(* IEC 61131-3 sources: plc-vscode/tests/st/test-ready/rusty/tests/lit/single/builtin, 5 files *)

(* ---- adr_ptr_arith_runtime.st ---- *)
// RUN: (%COMPILE %s && %RUN) | %CHECK %s
//
// `ADR(x) + N` is byte-stride pointer arithmetic — `ADR` is declared to
// return LWORD, so the `+` flows through the integer-arithmetic path; the
// receiver pointer ends up `N` bytes past the operand. Regression for #1749
// (previously panicked in `create_llvm_int_binary_expression`).

FUNCTION main
VAR
    arr : ARRAY[0..7] OF BYTE := [0, 0, 0, 0, 0, 0, 0, 0];
    pt  : REF_TO BYTE;
END_VAR

pt := ADR(arr) + 4;
pt^ := BYTE#16#AB;

// CHECK: arr[4]=171
printf('arr[4]=%d$N', arr[4]);

pt := ADR(arr) + 7;
pt^ := BYTE#16#5C;

// CHECK: arr[7]=92
printf('arr[7]=%d$N', arr[7]);

// Subtraction flows through the same path: take a pointer past the end
// and walk back. Writing to arr[2] via `ADR(arr[6]) - 4`.
pt := ADR(arr[6]) - 4;
pt^ := BYTE#16#11;

// CHECK: arr[2]=17
printf('arr[2]=%d$N', arr[2]);
END_FUNCTION

(* ---- shl_and_shr_must_cast_left_and_right_correctly.st ---- *)
// RUN: (%COMPILE %s && %RUN) | %CHECK %s

// SHL and SHR must cast left and right correctly
FUNCTION main
VAR
    value : BYTE;
END_VAR

value := BIT_LOAD_B2(BYTE#255, TRUE, 2, 2);

// CHECK: 255
printf('%d$N', value);

value := BIT_LOAD_B2(BYTE#255, FALSE, 2, 2);

// CHECK: 243
printf('%d$N', value);

END_FUNCTION

FUNCTION BIT_LOAD_B2 : BYTE
VAR_INPUT
	I : BYTE;
	D : BOOL;
	P : INT;
	N : INT;
END_VAR
VAR
    result : BYTE;
END_VAR

IF D THEN
	BIT_LOAD_B2 := ROL(SHR(BYTE#255, 8 - N) OR ROR(I, P), P);
ELSE
	BIT_LOAD_B2 := ROL(SHL(BYTE#255, N) AND ROR(I, P), P);
END_IF;

END_FUNCTION

(* ---- shl_must_be_usable_with_integers.st ---- *)
// RUN: (%COMPILE %s && %RUN) | %CHECK %s

// SHL must be usable with integers
FUNCTION main
VAR
    a : INT;
END_VAR
a := SHL(21,2);

// CHECK: 84
printf('%d$N', a);
END_FUNCTION

(* ---- shr_must_be_usable_with_integers.st ---- *)
// RUN: (%COMPILE %s && %RUN) | %CHECK %s

// SHR must be usable with integers
FUNCTION main
VAR
    a : INT;
END_VAR
a := SHR(21,2);

// CHECK: 5
printf('%d$N', a);
END_FUNCTION

(* ---- shr_unsigned_byte_logical_shift.st ---- *)
// RUN: (%COMPILE %s && %RUN) | %CHECK %s

// SHR on unsigned BYTE must use logical shift (zero-fill), not arithmetic shift
FUNCTION main
VAR
    b : BYTE;
    s : SINT;
END_VAR
b := SHR(BYTE#251, SINT#1);

// CHECK: 125
printf('%d$N', b);

s := SHR(SINT#-4, SINT#1);

// CHECK: -2
printf('%d$N', s);
END_FUNCTION
